SUBAPPLICATION Uebung_OPC_L01_AX (* Wie Training_01 (test_VV), aber lokal auf einem Geraet: Input_I1 schreibt per lokalem PUBLISH, Output_Q1 liest per lokalem SUBSCRIBE *)
  (* Standard: 61499-2; Description: Copyright (c) 2026 Meisterschulen am Ostbahnhof This program and the accompanying materials are made available under the terms of the Eclipse Public License 2.0 which is available at https://www.eclipse.org/legal/epl-2.0/ SPDX-License-Identifier: EPL-2.0 *)
  (* Version 1.0, 2026-10-18, Franz Höpfinger, Meisterschulen am Ostbahnhof, OPC-UA lokal auf einem Geraet (Meins/04_OPC_UA) *)
  PACKAGE Meins::OPC_UA_Lokal;
  IMPORT Meins::OPC_UA_Lokal::const::OpcUaLokal::L01_Q1_WRITE;
  IMPORT Meins::OPC_UA_Lokal::const::OpcUaLokal::L01_Q1_READ;
  IMPORT logiBUS::io::DI::logiBUS_DI::Input_I1;
  IMPORT logiBUS::io::DQ::logiBUS_DO::Output_Q1;
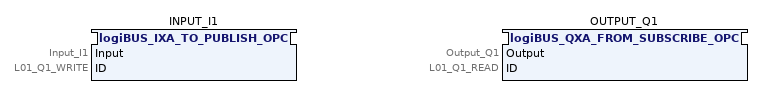
  SUBAPPS
    INPUT_I1 : MyLib::sys::logiBUS_IXA_TO_PUBLISH_OPC(Input := Input_I1, ID := L01_Q1_WRITE);
    OUTPUT_Q1 : MyLib::sys::logiBUS_QXA_FROM_SUBSCRIBE_OPC(Output := Output_Q1, ID := L01_Q1_READ);
  END_SUBAPPS
END_SUBAPPLICATION
